// TIA Portal V20 export
DATA_BLOCK "HMI_Statistik"   // DB2002
{ S7_Optimized_Access := 'FALSE' }
// stored: AutoNumber false
   VAR RETAIN
      Auftragsmenge : DInt := 0;
      Verpackungsmenge : DInt := 0;
      Verpackungszähler : DInt := 0;
      Beutelmenge : DInt := 0;
      "Letzte Zykluszeit" : Time := T#0MS;
      NIO_Behälter1 : DInt := 0;
      NIO_Behälter2 : DInt := 0;
      NIO_Behälter3 : DInt := 0;
      NIO_Behälter4 : DInt := 0;
      NIO_Behälter5 : DInt := 0;
      NIO_Behälter6 : DInt := 0;
      NIO_Behälter7 : DInt := 0;
      NIO_Behälter8 : DInt := 0;
      IO_Behälter1 : DInt := 0;
      IO_Behälter2 : DInt := 0;
      IO_Behälter3 : DInt := 0;
      IO_Behälter4 : DInt := 1000;
      IO_Behälter5 : DInt := 1000;
      NIO_BehälterMAX : DInt := 100;
      IO_BehälterMAX : DInt := 1000;
      Verpackungszähler_1 : DInt := 0;
      "Letzte Zykluszeit_POS_3_0" : Time := T#15S_228MS;
      "Letzte Zykluszeit_POS_3_0_in_s" : Real;
      "Durchschnitt Zykluszeit_POS_3_0" : Real;
      Restlaufzeit_POS_3_0 : Real;
      Zykluszeit_POS_3_0_in_s : Array[0..10] of Real;
      "Zaehler Alle Teile" : "HMI_Zaehler";
      "Zaehler IO Teile" : "HMI_Zaehler";
      "Zaehler NIO Teile" : "HMI_Zaehler";
      "IO 1" : "HMI_Zaehler";
      "IO 2" : "HMI_Zaehler";
      "IO 3" : "HMI_Zaehler";
      "IO 4" : "HMI_Zaehler";
      "IO 5" : "HMI_Zaehler";
      "NIO 1" { S7_SetPoint := 'True'} : "HMI_Zaehler";
      "NIO 2" { S7_SetPoint := 'True'} : "HMI_Zaehler";
      "NIO 3" { S7_SetPoint := 'True'} : "HMI_Zaehler";
      "NIO 4" { S7_SetPoint := 'True'} : "HMI_Zaehler";
      "NIO 5" { S7_SetPoint := 'True'} : "HMI_Zaehler";
      "NIO 6" { S7_SetPoint := 'True'} : "HMI_Zaehler";
   END_VAR
BEGIN
   "Zaehler Alle Teile".Schichtzaehler := 0;
   "Zaehler Alle Teile".Auftragszaehler := 0;
   "Zaehler Alle Teile".Gesamtzaehler := 0;
   "Zaehler IO Teile".Schichtzaehler := 0;
   "Zaehler IO Teile".Auftragszaehler := 0;
   "Zaehler IO Teile".Gesamtzaehler := 0;
   "Zaehler NIO Teile".Schichtzaehler := 0;
   "Zaehler NIO Teile".Auftragszaehler := 0;
   "Zaehler NIO Teile".Gesamtzaehler := 0;
   "IO 1".Schichtzaehler := 0;
   "IO 1".Auftragszaehler := 0;
   "IO 1".Gesamtzaehler := 0;
   "IO 2".Schichtzaehler := 0;
   "IO 2".Auftragszaehler := 0;
   "IO 2".Gesamtzaehler := 0;
   "IO 3".Schichtzaehler := 0;
   "IO 3".Auftragszaehler := 0;
   "IO 3".Gesamtzaehler := 0;
   "IO 4".Schichtzaehler := 0;
   "IO 4".Auftragszaehler := 0;
   "IO 4".Gesamtzaehler := 0;
   "IO 5".Schichtzaehler := 0;
   "IO 5".Auftragszaehler := 0;
   "IO 5".Gesamtzaehler := 0;
END_DATA_BLOCK
